// TIA Portal project "Project2" (V18)

(* hardware
DEVICE "S7-1500/ET200MP station_1"  S7-1500 station
   slot 0: "Rail_0"  Rack  6ES7 590-1***0-0AA0
   slot 1: "PLC_1"  CPU 1516-3 PN/DP  6ES7 516-3AN01-0AB0  V2.8
      slot 3: "CPU display_1"  6ES7591-1BA00-0AA0
      slot 32768: "PROFINET interface_1"  X1
         slot 32769: "Port_1"  X1 P1
         slot 32770: "Port_2"  X1 P2
      slot 33024: "PROFINET interface_2"  X2
         slot 33025: "Port_1"  X2 P1
      slot 33280: "DP interface_1"  X3
      slot 34817: "Virtual CP interface port_1"  Virtual CP interface port  Virtual CP interface port
DEVICE "GSD device_1"  GSD.Device.PN
   slot 0: "Rack"  Rack  V1.0
   slot 0: "IND360"  IND360 2 Block Format  MT-IND36XXXXXX  V1.0.0
      slot 0: "DAP 2 Block Parameter"  DAP 2 Block Parameter
      slot 1: "PROFINET"  PROFINET
         slot 1: "Port 1"  Port 1
         slot 2: "Port 2"  Port 2
      slot 1: "Measuring Block 1_1"  Measuring Block 1
         slot 0: "Parameter Access Point"  Parameter Access Point
         slot 1: "MB Command Value"  MB Command Value
         slot 2: "MB Channel Mask"  MB Channel Mask
         slot 3: "MB Command"  MB Command
         slot 4: "MB Measuring Value"  MB Measuring Value
         slot 5: "MB Device Status"  MB Device Status
         slot 6: "MB Response"  MB Response
      slot 2: "Status Block_1"  Status Block
         slot 0: "Parameter Access Point"  Parameter Access Point
         slot 1: "SB Reserved 1"  SB Reserved 1
         slot 2: "SB Reserved 2"  SB Reserved 2
         slot 3: "SB Reserved 3"  SB Reserved 3
         slot 4: "SB Command"  SB Command
         slot 5: "SB Status Group 1"  SB Status Group 1
         slot 6: "SB Status Group 2"  SB Status Group 2
         slot 7: "SB Status Group 3"  SB Status Group 3
         slot 8: "SB Response"  SB Response
DEVICE "HMI_1"  KTP400 Basic PN
   slot 0: "HMI_1"  KTP400 Basic PN  6AV2 123-2DB03-0AX0  17.0.0.0
   slot 1: "HMI_RT_1"  KTP400 Basic PN  6AV2 123-2DB03-0AX0  17.0.0.0
   slot 5: "HMI_1.IE_CP_1"  PROFINET Interface  17.0.0.0
      slot 1: "PROFINET Interface_1"  PROFINET Interface
         slot 1: "Port_1"  Port
*)

// ===== PLC "PLC_1"  CPU 1516-3 PN/DP =====

VAR_GLOBAL   // PLC tag table "Default tag table"
   "FirstScan" AT %M1.0 : Bool;
END_VAR

VAR_GLOBAL   // PLC tag table "IND"
   "T_MB_CmdValue" AT %QD0 : Real;
   "T_MB_Command" AT %QW6 : Word;
   "T_MB_Response" AT %IW6 : Word;
   "T_MB_Value" AT %ID0 : Real;
   "T_MB_DevStatus" AT %IW4 : Word;
   "T_SB_StaGroup1" AT %IW8 : Word;
   "T_SB_StaGroup2" AT %IW10 : Word;
   "T_SB_StaGroup3" AT %IW12 : Word;
   "T_SB_Response" AT %IW14 : Word;
   "T_SB_Command" AT %QW14 : Word;
   "AlibiGross_Byte(0)" AT %MB50 : Byte;
   "AlibiGross_Byte(1)" AT %MB51 : Byte;
   "AlibiGross_Byte(2)" AT %MB52 : Byte;
   "AlibiGross_Byte(3)" AT %MB53 : Byte;
   "AlibiNet_Byte(0)" AT %MB58 : Byte;
   "AlibiNet_Byte(1)" AT %MB59 : Byte;
   "AlibiNet_Byte(2)" AT %MB60 : Byte;
   "AlibiNet_Byte(3)" AT %MB61 : Byte;
   "AlibiTare_Byte(0)" AT %MB66 : Byte;
   "AlibiTare_Byte(1)" AT %MB67 : Byte;
   "AlibiTare_Byte(2)" AT %MB68 : Byte;
   "AlibiTare_Byte(3)" AT %MB69 : Byte;
   "AlibiGross_Real" AT %MD50 : Real;
   "AlibiNet_Real" AT %MD58 : Real;
   "AlibiTare_Real" AT %MD66 : Real;
END_VAR

TYPE "SAI_MB_DeviceStatus"
VERSION : 0.1
   STRUCT
      "Alternate weight unit" : Bool;
      "Run flat" : Bool;
      "Device specific bit 2" : Bool;
      "Device specific bit 3" : Bool;
      "Device specific bit 4" : Bool;
      "Device specific bit 5" : Bool;
      "Device specific bit 6" : Bool;
      "Device specific bit 7" : Bool;
      "Sequence bit 0" : Bool;
      "Sequence bit 1" : Bool;
      "Heart Beat" : Bool;
      "Data OK" : Bool;
      "Alarm Condition" : Bool;
      "Center of Zero" : Bool;
      Motion : Bool;
      "Net Mode" : Bool;
   END_STRUCT;
END_TYPE

TYPE "SAI_SB_RedAlert"
   STRUCT
      "Zero out of range" : Bool;
      "Symetry errors" : Bool;
      "LC Temperature out of normal temperature" : Bool;
      "Weights and measures failure" : Bool;
      "Foreign device detected" : Bool;
      "Test mode" : Bool;
      "LC temperature out of operatio" : Bool;
      "LC parameters block checksum error" : Bool;
      "Calibration error" : Bool;
      "Out of A/D range over/under" : Bool;
      "Checksu failure" : Bool;
      "Weight blocked" : Bool;
      "LC Missing" : Bool;
      "Customer-defined overload" : Bool;
      "Customer-defined underload" : Bool;
   END_STRUCT;
END_TYPE

TYPE "SAI_SB_Alarm"
   STRUCT
      "LC overload in operation range" : Bool;
      "LC Mix" : Bool;
      "Application defined 1" : Bool;
      "Application defined 2" : Bool;
      "Application defined 3" : Bool;
      "Application defined 4" : Bool;
      "Application defined 5" : Bool;
      "Application defined 7" : Bool;
      "Rate of change error" : Bool;
      "Communication error" : Bool;
      "Over / under voltage" : Bool;
      "Weight drift" : Bool;
      Breach : Bool;
      "Calibration expired" : Bool;
      "Over Current" : Bool;
      "LC overload in normal range" : Bool;
   END_STRUCT;
END_TYPE

DATA_BLOCK "SAI_Cyclic_CheckAlive_DB"   // DB1
{ S7_Optimized_Access := 'FALSE' }
VERSION : 0.1
// stored: InstanceOfName SAI_Cyclic_CheckAlive
"SAI_Cyclic_CheckAlive"
BEGIN
END_DATA_BLOCK

DATA_BLOCK "SAI_Cyclic_WeightProc_DB"   // DB2
{ S7_Optimized_Access := 'FALSE' }
VERSION : 0.1
// stored: InstanceOfName SAI_Cyclic_WeightProc
"SAI_Cyclic_WeightProc"
BEGIN
END_DATA_BLOCK

FUNCTION_BLOCK "SAI_Cyclic_CheckAlive"   // FB1, LAD
TITLE = Check HearBeat status bit and update the Alive bit
{ S7_Optimized_Access := 'FALSE' }
VERSION : 0.1
   VAR_INPUT
      MB_DevStatus : Word;
   END_VAR
   VAR_OUTPUT
      Alive : Bool;
      HeartBeat : Bool;
   END_VAR
   VAR
      PTrigHeart : Bool;
      NTrigHeart : Bool;
      bResetTimer : Bool;
      IEC_Timer : IEC_TIMER;
   END_VAR
   VAR_TEMP
      DevStatus : "SAI_MB_DeviceStatus";
   END_VAR
   VAR_TEMP   // added for the SCL form of the ladder/FBD networks
      _w1 : Bool;
      _w2 : Bool;
      _w3 : Bool;
   END_VAR
BEGIN

REGION Network 1: 复制设备状态到结构体 / Gets the cyclic device status - HeartBeat bit
   // Gets the cyclic device status - HeartBeat bit
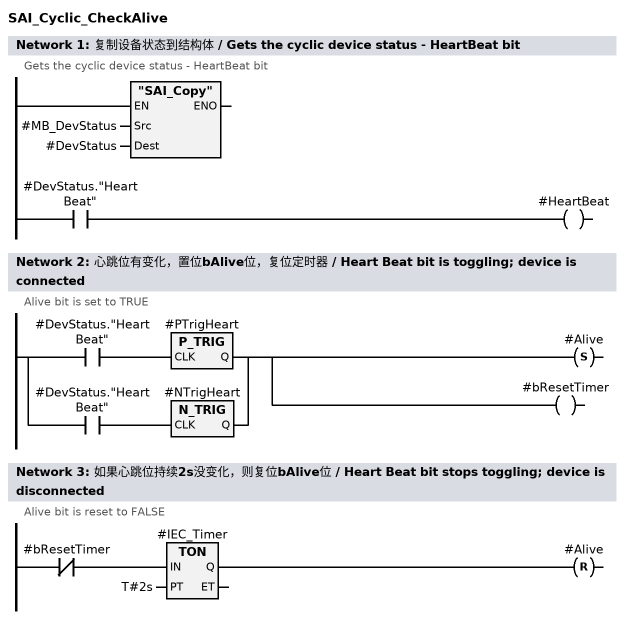
   RUNG wire#powerrail
      "SAI_Copy"(Src := #MB_DevStatus, Dest := #DevStatus)
   END_RUNG
   RUNG wire#powerrail
      Contact( #DevStatus."Heart Beat" )
      Coil( #HeartBeat )
   END_RUNG
   // the same network as SCL:
   "SAI_Copy"(Src := #MB_DevStatus, Dest := #DevStatus);
   #HeartBeat := #DevStatus."Heart Beat";
END_REGION

REGION Network 2: 心跳位有变化，置位bAlive位，复位定时器 / Heart Beat bit is toggling; device is connected
   // Alive bit is set to TRUE
   RUNG wire#powerrail
      Contact( #DevStatus."Heart Beat" )
      P_Trig( #PTrigHeart )
      wire#w1
      S_Coil( #Alive )
   END_RUNG
   RUNG wire#powerrail
      Contact( #DevStatus."Heart Beat" )
      N_Trig( #NTrigHeart )
   END_RUNG wire#w1
   RUNG wire#w1
      Coil( #bResetTimer )
   END_RUNG
   // the same network as SCL:
   #_w1 := #DevStatus."Heart Beat" AND NOT #PTrigHeart;   // rising edge
   #PTrigHeart := #DevStatus."Heart Beat";
   #_w2 := NOT #DevStatus."Heart Beat" AND #NTrigHeart;   // falling edge
   #NTrigHeart := #DevStatus."Heart Beat";
   #_w3 := #_w1 OR #_w2;
   IF #_w3 THEN #Alive := TRUE; END_IF;
   #bResetTimer := #_w3;
END_REGION

REGION Network 3: 如果心跳位持续2s没变化，则复位bAlive位 / Heart Beat bit stops toggling; device is disconnected
   // Alive bit is reset to FALSE
   #IEC_Timer.TON(IN := NOT #bResetTimer, PT := T#2s);
   IF #IEC_Timer.Q THEN #Alive := FALSE; END_IF;
END_REGION
END_FUNCTION_BLOCK

FUNCTION_BLOCK "SAI_Cyclic_WeightProc"   // FB2, LAD
TITLE = Cyclic Weighing Process: Send PLC commands and read Weight data and device status bits
{ S7_Optimized_Access := 'FALSE' }
VERSION : 0.1
   VAR_INPUT
      WeightCmd : Word := 3;
      MB_DevStatus : Word;
   END_VAR
   VAR_OUTPUT
      RealTimeWeight : Real;
      StableWeight : Real;
      DataOK : Bool;
      Motion : Bool;
      NetMode : Bool;
      Alarm : Bool;
      Done : Bool;
      Error : Bool;
   END_VAR
   VAR_IN_OUT
      TareImmediate : Bool;
      TareStable : Bool;
      ZeroImmediate : Bool;
      ZeroStable : Bool;
      PreTareValue : Real;
      PreTare : Bool;
      ClearTare : Bool;
      MB_Value : Real;
      MB_Response : Word;
      MB_CmdValue : Real;
      MB_Command : Word;
   END_VAR
   VAR
      WriteTrigger : Bool;
      RestoreTrigger : Bool;
      Cmd : Int;
      TareStablePTrigger : Bool;
      ZeroStablePTrigger : Bool;
      ZeroImmedTrigger : Bool;
      TareImmedTrigger : Bool;
      ClearTareTrigger : Bool;
      PreTareTrigger : Bool;
   END_VAR
   VAR_TEMP
      DevStatus : "SAI_MB_DeviceStatus";
   END_VAR
   VAR_TEMP   // added for the SCL form of the ladder/FBD networks
      _w1 : Bool;
   END_VAR
BEGIN

REGION Network 1: 第一次运行时，将默认重量命令赋值给循环区命令 / During 1st PLC scan, moves the default weight reporting command to the cyclic command output word
   // 第一次扫描，写入重量命令 / During 1st scan, moves the default weight reporting command to the cyclic command output word
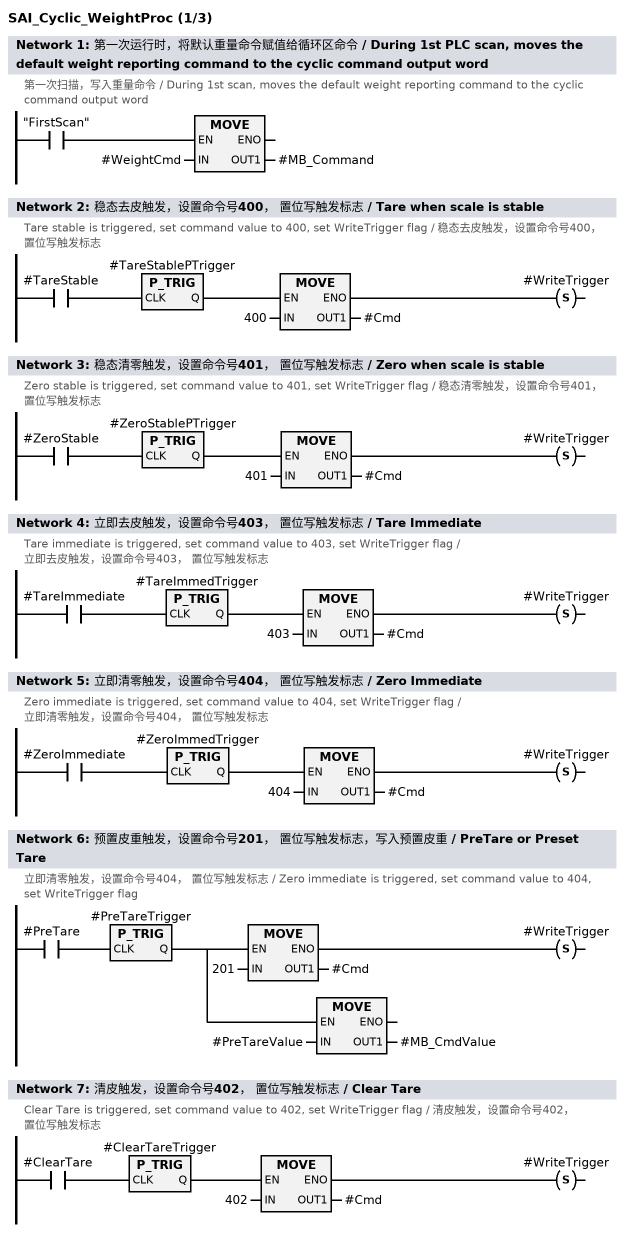
   RUNG wire#powerrail
      Contact( "FirstScan" )
      { S7_GenerateENO := "TRUE" } Move(in := #WeightCmd, out1 => #MB_Command)
   END_RUNG
   // the same network as SCL:
   IF "FirstScan" THEN #MB_Command := #WeightCmd; END_IF;
END_REGION

REGION Network 2: 稳态去皮触发，设置命令号400， 置位写触发标志 / Tare when scale is stable
   // Tare stable is triggered, set command value to 400, set WriteTrigger flag / 稳态去皮触发，设置命令号400， 置位写触发标志
   RUNG wire#powerrail
      Contact( #TareStable )
      P_Trig( #TareStablePTrigger )
      { S7_GenerateENO := "TRUE" } Move(in := 400, out1 => #Cmd)
      S_Coil( #WriteTrigger )
   END_RUNG
   // the same network as SCL:
   // ENO of a box is taken as its EN; it also drops when the box reports an error
   #_w1 := #TareStable AND NOT #TareStablePTrigger;   // rising edge
   #TareStablePTrigger := #TareStable;
   IF #_w1 THEN
       #Cmd := 400;
       #WriteTrigger := TRUE;
   END_IF;
END_REGION

REGION Network 3: 稳态清零触发，设置命令号401， 置位写触发标志 / Zero when scale is stable
   // Zero stable is triggered, set command value to 401, set WriteTrigger flag / 稳态清零触发，设置命令号401， 置位写触发标志
   RUNG wire#powerrail
      Contact( #ZeroStable )
      P_Trig( #ZeroStablePTrigger )
      { S7_GenerateENO := "TRUE" } Move(in := 401, out1 => #Cmd)
      S_Coil( #WriteTrigger )
   END_RUNG
   // the same network as SCL:
   // ENO of a box is taken as its EN; it also drops when the box reports an error
   #_w1 := #ZeroStable AND NOT #ZeroStablePTrigger;   // rising edge
   #ZeroStablePTrigger := #ZeroStable;
   IF #_w1 THEN
       #Cmd := 401;
       #WriteTrigger := TRUE;
   END_IF;
END_REGION

REGION Network 4: 立即去皮触发，设置命令号403， 置位写触发标志 / Tare Immediate
   // Tare immediate is triggered, set command value to 403, set WriteTrigger flag / 立即去皮触发，设置命令号403， 置位写触发标志
   RUNG wire#powerrail
      Contact( #TareImmediate )
      P_Trig( #TareImmedTrigger )
      { S7_GenerateENO := "TRUE" } Move(in := 403, out1 => #Cmd)
      S_Coil( #WriteTrigger )
   END_RUNG
   // the same network as SCL:
   // ENO of a box is taken as its EN; it also drops when the box reports an error
   #_w1 := #TareImmediate AND NOT #TareImmedTrigger;   // rising edge
   #TareImmedTrigger := #TareImmediate;
   IF #_w1 THEN
       #Cmd := 403;
       #WriteTrigger := TRUE;
   END_IF;
END_REGION

REGION Network 5: 立即清零触发，设置命令号404， 置位写触发标志 / Zero Immediate
   // Zero immediate is triggered, set command value to 404, set WriteTrigger flag / 立即清零触发，设置命令号404， 置位写触发标志
   RUNG wire#powerrail
      Contact( #ZeroImmediate )
      P_Trig( #ZeroImmedTrigger )
      { S7_GenerateENO := "TRUE" } Move(in := 404, out1 => #Cmd)
      S_Coil( #WriteTrigger )
   END_RUNG
   // the same network as SCL:
   // ENO of a box is taken as its EN; it also drops when the box reports an error
   #_w1 := #ZeroImmediate AND NOT #ZeroImmedTrigger;   // rising edge
   #ZeroImmedTrigger := #ZeroImmediate;
   IF #_w1 THEN
       #Cmd := 404;
       #WriteTrigger := TRUE;
   END_IF;
END_REGION

REGION Network 6: 预置皮重触发，设置命令号201， 置位写触发标志，写入预置皮重 / PreTare or Preset Tare
   // 立即清零触发，设置命令号404， 置位写触发标志 / Zero immediate is triggered, set command value to 404, set WriteTrigger flag
   RUNG wire#powerrail
      Contact( #PreTare )
      P_Trig( #PreTareTrigger )
      wire#w1
      { S7_GenerateENO := "TRUE" } Move(in := 201, out1 => #Cmd)
      S_Coil( #WriteTrigger )
   END_RUNG
   RUNG wire#w1
      { S7_GenerateENO := "TRUE" } Move(in := #PreTareValue, out1 => #MB_CmdValue)
   END_RUNG
   // the same network as SCL:
   // ENO of a box is taken as its EN; it also drops when the box reports an error
   #_w1 := #PreTare AND NOT #PreTareTrigger;   // rising edge
   #PreTareTrigger := #PreTare;
   IF #_w1 THEN
       #Cmd := 201;
       #WriteTrigger := TRUE;
       #MB_CmdValue := #PreTareValue;
   END_IF;
END_REGION

REGION Network 7: 清皮触发，设置命令号402， 置位写触发标志 / Clear Tare
   // Clear Tare is triggered, set command value to 402, set WriteTrigger flag / 清皮触发，设置命令号402， 置位写触发标志
   RUNG wire#powerrail
      Contact( #ClearTare )
      P_Trig( #ClearTareTrigger )
      { S7_GenerateENO := "TRUE" } Move(in := 402, out1 => #Cmd)
      S_Coil( #WriteTrigger )
   END_RUNG
   // the same network as SCL:
   // ENO of a box is taken as its EN; it also drops when the box reports an error
   #_w1 := #ClearTare AND NOT #ClearTareTrigger;   // rising edge
   #ClearTareTrigger := #ClearTare;
   IF #_w1 THEN
       #Cmd := 402;
       #WriteTrigger := TRUE;
   END_IF;
END_REGION

REGION Network 8: 将命令值赋值给输出循环区，复位标志，清除命令值 / Deliver the command
   // Move the command value to output, reset flags / 将命令输出，置位标志
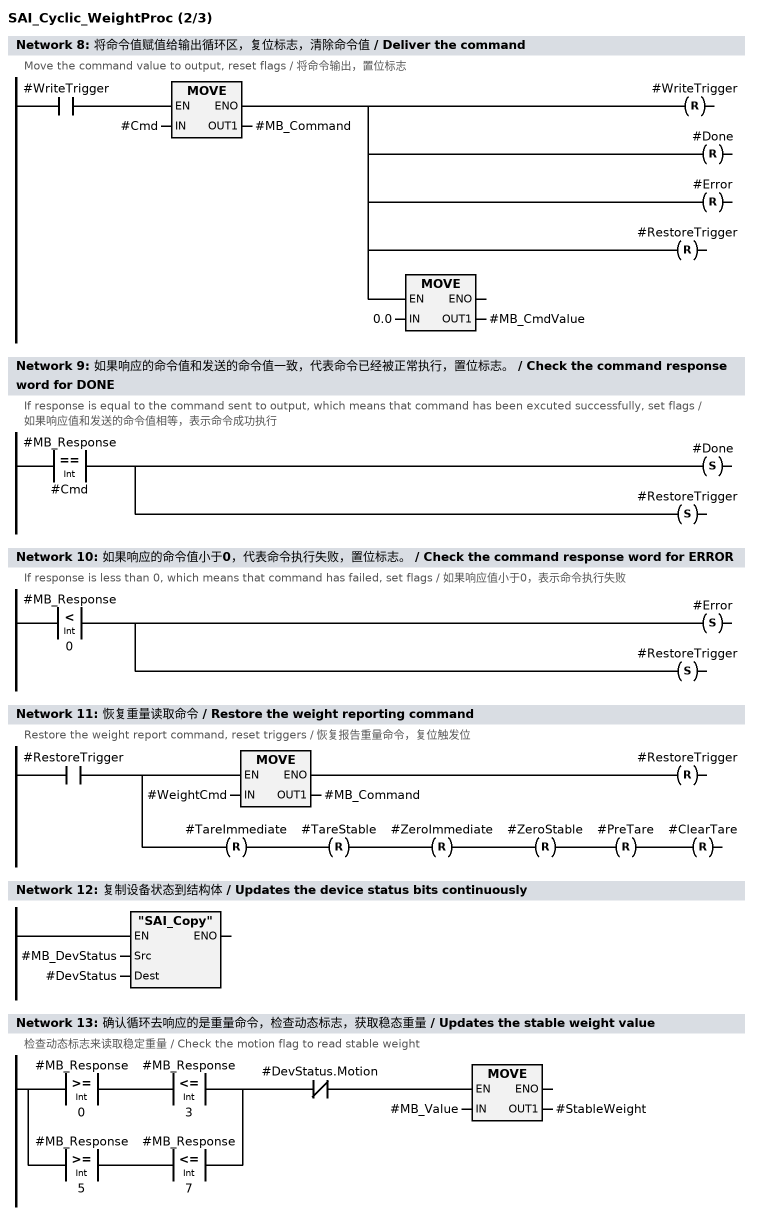
   RUNG wire#powerrail
      Contact( #WriteTrigger )
      { S7_GenerateENO := "TRUE" } Move(in := #Cmd, out1 => #MB_Command)
      wire#w1
      R_Coil( #WriteTrigger )
   END_RUNG
   RUNG wire#w1
      R_Coil( #Done )
   END_RUNG
   RUNG wire#w1
      R_Coil( #Error )
   END_RUNG
   RUNG wire#w1
      R_Coil( #RestoreTrigger )
   END_RUNG
   RUNG wire#w1
      { S7_GenerateENO := "TRUE" } Move(in := 0.0, out1 => #MB_CmdValue)
   END_RUNG
   // the same network as SCL:
   // ENO of a box is taken as its EN; it also drops when the box reports an error
   IF #WriteTrigger THEN #MB_Command := #Cmd; END_IF;
   #_w1 := #WriteTrigger;
   IF #_w1 THEN
       #WriteTrigger := FALSE;
       #Done := FALSE;
       #Error := FALSE;
       #RestoreTrigger := FALSE;
       #MB_CmdValue := 0.0;
   END_IF;
END_REGION

REGION Network 9: 如果响应的命令值和发送的命令值一致，代表命令已经被正常执行，置位标志。 / Check the command response word for DONE
   // If response is equal to the command sent to output, which means that command has been excuted successfully, set flags / 如果响应值和发送的命令值相等，表示命令成功执行
   RUNG wire#powerrail
      { S7_Templates := "SrcType := Int" } EQ_Contact(in1 := #MB_Response, in2 := #Cmd)
      wire#w1
      S_Coil( #Done )
   END_RUNG
   RUNG wire#w1
      S_Coil( #RestoreTrigger )
   END_RUNG
   // the same network as SCL:
   IF #MB_Response = #Cmd THEN
       #Done := TRUE;
       #RestoreTrigger := TRUE;
   END_IF;
END_REGION

REGION Network 10: 如果响应的命令值小于0，代表命令执行失败，置位标志。 / Check the command response word for ERROR
   // If response is less than 0, which means that command has failed, set flags / 如果响应值小于0，表示命令执行失败
   RUNG wire#powerrail
      { S7_Templates := "SrcType := Int" } LT_Contact(in1 := #MB_Response, in2 := 0)
      wire#w1
      S_Coil( #Error )
   END_RUNG
   RUNG wire#w1
      S_Coil( #RestoreTrigger )
   END_RUNG
   // the same network as SCL:
   IF #MB_Response < 0 THEN
       #Error := TRUE;
       #RestoreTrigger := TRUE;
   END_IF;
END_REGION

REGION Network 11: 恢复重量读取命令 / Restore the weight reporting command
   // Restore the weight report command, reset triggers / 恢复报告重量命令，复位触发位
   RUNG wire#powerrail
      Contact( #RestoreTrigger )
      wire#w1
      { S7_GenerateENO := "TRUE" } Move(in := #WeightCmd, out1 => #MB_Command)
      R_Coil( #RestoreTrigger )
   END_RUNG
   RUNG wire#w1
      R_Coil( #TareImmediate )
      R_Coil( #TareStable )
      R_Coil( #ZeroImmediate )
      R_Coil( #ZeroStable )
      R_Coil( #PreTare )
      R_Coil( #ClearTare )
   END_RUNG
   // the same network as SCL:
   // ENO of a box is taken as its EN; it also drops when the box reports an error
   IF #RestoreTrigger THEN #MB_Command := #WeightCmd; END_IF;
   #_w1 := #RestoreTrigger;
   IF #_w1 THEN
       #RestoreTrigger := FALSE;
       #TareImmediate := FALSE;
       #TareStable := FALSE;
       #ZeroImmediate := FALSE;
       #ZeroStable := FALSE;
       #PreTare := FALSE;
       #ClearTare := FALSE;
   END_IF;
END_REGION

REGION Network 12: 复制设备状态到结构体 / Updates the device status bits continuously
   RUNG wire#powerrail
      "SAI_Copy"(Src := #MB_DevStatus, Dest := #DevStatus)
   END_RUNG
   // the same network as SCL:
   "SAI_Copy"(Src := #MB_DevStatus, Dest := #DevStatus);
END_REGION

REGION Network 13: 确认循环去响应的是重量命令，检查动态标志，获取稳态重量 / Updates the stable weight value
   // 检查动态标志来读取稳定重量 / Check the motion flag to read stable weight
   RUNG wire#powerrail
      { S7_Templates := "SrcType := Int" } GE_Contact(in1 := #MB_Response, in2 := 0)
      { S7_Templates := "SrcType := Int" } LE_Contact(in1 := #MB_Response, in2 := 3)
      wire#w1
      I_Contact( #DevStatus.Motion )
      { S7_GenerateENO := "TRUE" } Move(in := #MB_Value, out1 => #StableWeight)
   END_RUNG
   RUNG wire#powerrail
      { S7_Templates := "SrcType := Int" } GE_Contact(in1 := #MB_Response, in2 := 5)
      { S7_Templates := "SrcType := Int" } LE_Contact(in1 := #MB_Response, in2 := 7)
   END_RUNG wire#w1
   // the same network as SCL:
   IF (((#MB_Response >= 0) AND (#MB_Response <= 3)) OR ((#MB_Response >= 5) AND (#MB_Response <= 7))) AND NOT #DevStatus.Motion THEN
       #StableWeight := #MB_Value;
   END_IF;
END_REGION

REGION Network 14: 确认循环去响应的是重量命令，读取实时的重量 / Updates the real time weight value
   // 读取实时重量 / Read real time weight
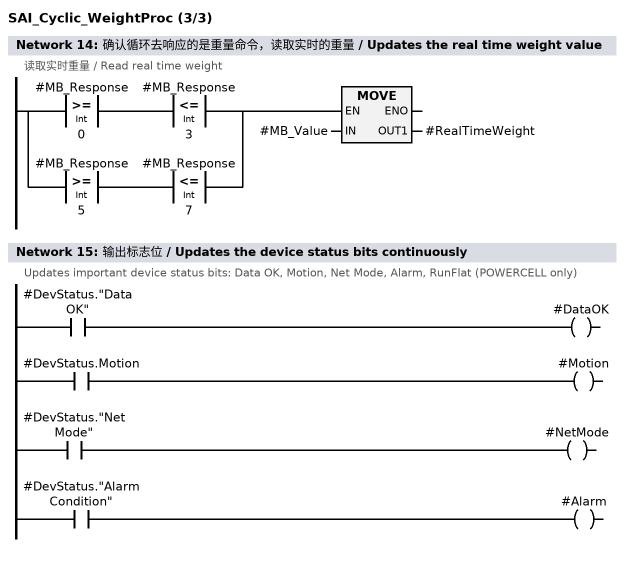
   RUNG wire#powerrail
      { S7_Templates := "SrcType := Int" } GE_Contact(in1 := #MB_Response, in2 := 0)
      { S7_Templates := "SrcType := Int" } LE_Contact(in1 := #MB_Response, in2 := 3)
      wire#w1
      { S7_GenerateENO := "TRUE" } Move(in := #MB_Value, out1 => #RealTimeWeight)
   END_RUNG
   RUNG wire#powerrail
      { S7_Templates := "SrcType := Int" } GE_Contact(in1 := #MB_Response, in2 := 5)
      { S7_Templates := "SrcType := Int" } LE_Contact(in1 := #MB_Response, in2 := 7)
   END_RUNG wire#w1
   // the same network as SCL:
   IF ((#MB_Response >= 0) AND (#MB_Response <= 3)) OR ((#MB_Response >= 5) AND (#MB_Response <= 7)) THEN
       #RealTimeWeight := #MB_Value;
   END_IF;
END_REGION

REGION Network 15: 输出标志位 / Updates the device status bits continuously
   // Updates important device status bits: Data OK, Motion, Net Mode, Alarm, RunFlat (POWERCELL only)
   RUNG wire#powerrail
      Contact( #DevStatus."Data OK" )
      Coil( #DataOK )
   END_RUNG
   RUNG wire#powerrail
      Contact( #DevStatus.Motion )
      Coil( #Motion )
   END_RUNG
   RUNG wire#powerrail
      Contact( #DevStatus."Net Mode" )
      Coil( #NetMode )
   END_RUNG
   RUNG wire#powerrail
      Contact( #DevStatus."Alarm Condition" )
      Coil( #Alarm )
   END_RUNG
   // the same network as SCL:
   #DataOK := #DevStatus."Data OK";
   #Motion := #DevStatus.Motion;
   #NetMode := #DevStatus."Net Mode";
   #Alarm := #DevStatus."Alarm Condition";
END_REGION
END_FUNCTION_BLOCK

FUNCTION "SAI_Copy" : Void   // FC1, LAD
{ S7_Optimized_Access := 'FALSE' }
VERSION : 0.1
   VAR_INPUT
      Src : Variant;
   END_VAR
   VAR_IN_OUT
      Dest : Variant;
   END_VAR
   VAR_TEMP
      TmpBuf : Array[0..100] of Byte;
      TmpRet : Int;
      TmpPos : DInt;
   END_VAR
BEGIN

REGION Network 1
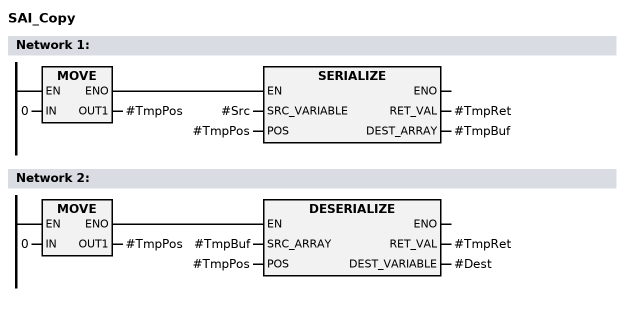
   // no SCL statement known for Serialize: written as a call
   #TmpPos := 0;
   #TmpRet := Serialize(SRC_VARIABLE := #Src, POS := #TmpPos, DEST_ARRAY => #TmpBuf);
END_REGION

REGION Network 2
   // no SCL statement known for Deserialize: written as a call
   #TmpPos := 0;
   #TmpRet := Deserialize(SRC_ARRAY := #TmpBuf, POS := #TmpPos, DEST_VARIABLE => #Dest);
END_REGION
END_FUNCTION

FUNCTION "MT_ACT_Application" : Void   // FC2, LAD
{ S7_Optimized_Access := 'FALSE' }
VERSION : 0.1
BEGIN

REGION Network 1: 循环重量处理 / Cyclic Weighing Data
   // 读取实时重量RealTimeWeight和稳态重量StableWeight，数据正常位DataOK，动态标志位Motion，净重模式位NetMode和警报位Alarm。
   // 上升沿触发执行稳态去皮TareStable，稳态清零ZeroStable，立即去皮TareImmediate，立即清零ZeroImmediate，预置皮重PreTare和清皮ClearTare，执行过程中，执行成功Done和失败Error的标志会复位为0，执行完成会置位Done或者Error来指示命令执行结果。清零去皮处理时，实时重量和稳态重量会保持不更新。
   // 在清零和去皮执行完成后，重量命令WeightCmd会自动发送一次，让MB Measuring Value循环区报告重量值，默认将恢复WeightCmd为读取净重（命令号3）。
   // 参照参数表中的重量命令值进行设置，执行清零或者去皮处理后，则会读取到对应的重量。
   // All the cyclical read and write commands can be issued from this Function Block.
   // The cyclic commands are triggered following a positive trigger. These commands are Tare Immediate, Tare Stable, Zero Immediate, Zero Stable, Pretare and Clear Tare. 
   // Upon successful execution of these commands, the DONE output bit will be set ON.
   // ERROR output bit will be set on if there is an error with the command execution.
   // Note: Only one cyclic command is possible at any one time.
   // If Net weight is required after executed a zero or tare command, insert decimal value "3" into the "WeightCmd" variable before triggering the cyclic scale command. Else, with decimal value "1" in the "WeightCmd" variable, the Function Block will return Gross Weight after the cyclic scale command. 
   // "DataOK" bit is set ON when the scale is in operation mode, not overloaded and not underload.
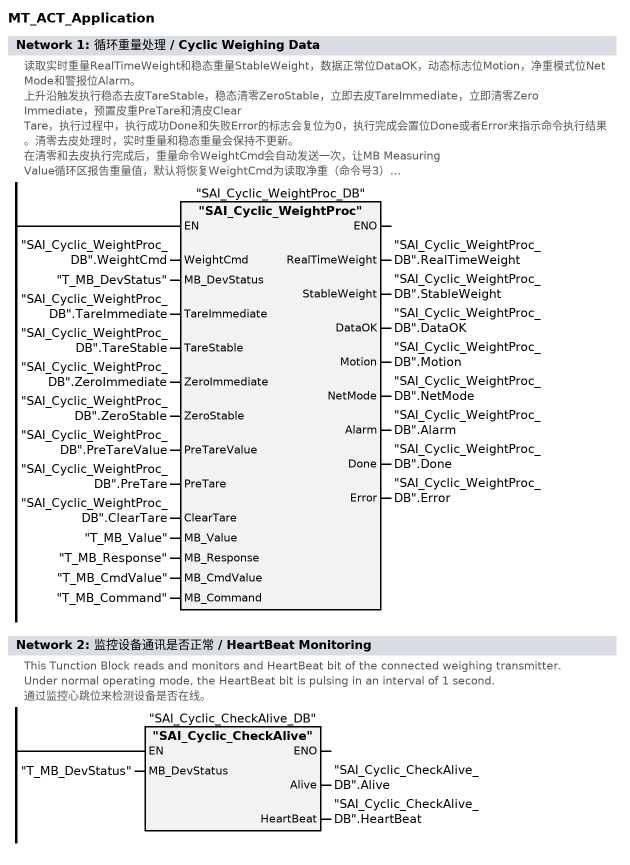
   RUNG wire#powerrail
      "SAI_Cyclic_WeightProc_DB"(WeightCmd := "SAI_Cyclic_WeightProc_DB".WeightCmd, MB_DevStatus := "T_MB_DevStatus", TareImmediate := "SAI_Cyclic_WeightProc_DB".TareImmediate, TareStable := "SAI_Cyclic_WeightProc_DB".TareStable, ZeroImmediate := "SAI_Cyclic_WeightProc_DB".ZeroImmediate, ZeroStable := "SAI_Cyclic_WeightProc_DB".ZeroStable, PreTareValue := "SAI_Cyclic_WeightProc_DB".PreTareValue, PreTare := "SAI_Cyclic_WeightProc_DB".PreTare, ClearTare := "SAI_Cyclic_WeightProc_DB".ClearTare, MB_Value := "T_MB_Value", MB_Response := "T_MB_Response", MB_CmdValue := "T_MB_CmdValue", MB_Command := "T_MB_Command", RealTimeWeight => "SAI_Cyclic_WeightProc_DB".RealTimeWeight, StableWeight => "SAI_Cyclic_WeightProc_DB".StableWeight, DataOK => "SAI_Cyclic_WeightProc_DB".DataOK, Motion => "SAI_Cyclic_WeightProc_DB".Motion, NetMode => "SAI_Cyclic_WeightProc_DB".NetMode, Alarm => "SAI_Cyclic_WeightProc_DB".Alarm, Done => "SAI_Cyclic_WeightProc_DB".Done, Error => "SAI_Cyclic_WeightProc_DB".Error)
   END_RUNG
   // the same network as SCL:
   "SAI_Cyclic_WeightProc_DB"(WeightCmd := "SAI_Cyclic_WeightProc_DB".WeightCmd,   // "SAI_Cyclic_WeightProc"
                           MB_DevStatus := "T_MB_DevStatus",
                           TareImmediate := "SAI_Cyclic_WeightProc_DB".TareImmediate,
                           TareStable := "SAI_Cyclic_WeightProc_DB".TareStable,
                           ZeroImmediate := "SAI_Cyclic_WeightProc_DB".ZeroImmediate,
                           ZeroStable := "SAI_Cyclic_WeightProc_DB".ZeroStable,
                           PreTareValue := "SAI_Cyclic_WeightProc_DB".PreTareValue,
                           PreTare := "SAI_Cyclic_WeightProc_DB".PreTare,
                           ClearTare := "SAI_Cyclic_WeightProc_DB".ClearTare,
                           MB_Value := "T_MB_Value",
                           MB_Response := "T_MB_Response",
                           MB_CmdValue := "T_MB_CmdValue",
                           MB_Command := "T_MB_Command",
                           RealTimeWeight => "SAI_Cyclic_WeightProc_DB".RealTimeWeight,
                           StableWeight => "SAI_Cyclic_WeightProc_DB".StableWeight,
                           DataOK => "SAI_Cyclic_WeightProc_DB".DataOK,
                           Motion => "SAI_Cyclic_WeightProc_DB".Motion,
                           NetMode => "SAI_Cyclic_WeightProc_DB".NetMode,
                           Alarm => "SAI_Cyclic_WeightProc_DB".Alarm,
                           Done => "SAI_Cyclic_WeightProc_DB".Done,
                           Error => "SAI_Cyclic_WeightProc_DB".Error);
END_REGION

REGION Network 2: 监控设备通讯是否正常 / HeartBeat Monitoring
   // This Tunction Block reads and monitors and HeartBeat bit of the connected weighing transmitter.
   // Under normal operating mode, the HeartBeat bit is pulsing in an interval of 1 second.
   // 通过监控心跳位来检测设备是否在线。
   RUNG wire#powerrail
      "SAI_Cyclic_CheckAlive_DB"(MB_DevStatus := "T_MB_DevStatus", Alive => "SAI_Cyclic_CheckAlive_DB".Alive, HeartBeat => "SAI_Cyclic_CheckAlive_DB".HeartBeat)
   END_RUNG
   // the same network as SCL:
   "SAI_Cyclic_CheckAlive_DB"(MB_DevStatus := "T_MB_DevStatus",   // "SAI_Cyclic_CheckAlive"
                           Alive => "SAI_Cyclic_CheckAlive_DB".Alive,
                           HeartBeat => "SAI_Cyclic_CheckAlive_DB".HeartBeat);
END_REGION
END_FUNCTION

ORGANIZATION_BLOCK "Main"   // OB1, LAD, ProgramCycle
TITLE = "Main Program Sweep (Cycle)"
{ S7_Optimized_Access := 'TRUE' }
VERSION : 0.1
   VAR_INPUT
      Initial_Call : Bool;   // Initial call of this OB
      Remanence : Bool;   // =True, if remanent data are available
   END_VAR
BEGIN

REGION Network 1
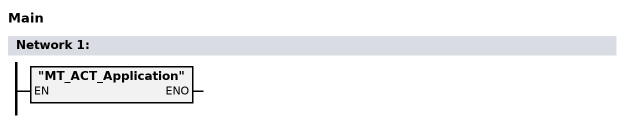
   RUNG wire#powerrail
      "MT_ACT_Application"()
   END_RUNG
   // the same network as SCL:
   "MT_ACT_Application"();
END_REGION
END_ORGANIZATION_BLOCK

(* ===== HMI "HMI_RT_1" =====
system functions are stored by id; their names below are inferred from use
connection "HMI_Connection_1": ETHERNET, SMART_S7_1500_OMS

HMI tags "Default tag table"
   "Tag_ScreenNumber" : UInt, internal
   "xHeartbeat" : Bool = PLC SAI_Cyclic_CheckAlive_DB.HeartBeat AT %DB1.DBX2.1, 1 s
   "rCurrentWeight" : Real = PLC SAI_Cyclic_WeightProc_DB.StableWeight AT %DB2.DBD8, 1 s
   "xZeroScale" : Bool = PLC SAI_Cyclic_WeightProc_DB.ZeroStable AT %DB2.DBX14.3, 1 s
   "xClearTare" : Bool = PLC SAI_Cyclic_WeightProc_DB.ClearTare AT %DB2.DBX20.1, 1 s
   "xSetTare" : Bool = PLC SAI_Cyclic_WeightProc_DB.TareStable AT %DB2.DBX14.1, 1 s

Template "Template_1" 480x272
   Button "Exit" at 388,227 size 63x44; TextOff 'Exit'; PictureOff "ExitRuntime_KTP400_Basic_PN_TR"; PictureOn "ExitRuntime_KTP400_Basic_PN_TR"
      on Release: StopRuntime(0)
   Button "Template_Button" at 268,227 size 63x44; TextOff 'Text'
   Button "Template_Button_1" at 148,227 size 63x44; TextOff 'Text'
   Button "Start screen" at 28,227 size 63x44; TextOff 'Start screen'; PictureOff "NavigateHome_KTP400_Basic_PN_TR"; PictureOn "NavigateHome_KTP400_Basic_PN_TR"
      on Release: ActivateScreen("Root screen", 0)
   SymbolicIOField "Symbolic_IO_Field_Screen" at 82,8 size 311x29; TextOff '0'; TextOn '1'; TextList "TextList_ScreenNames"
      ProcessValue <- "Tag_ScreenNumber"
      on Change: ActivateScreenByNumber("Tag_ScreenNumber", 0)
   DateTimeField "HmiScreenItemData" at 395,22 size 85x22
   DateTimeField "HmiScreenItemData_1" at 395,0 size 85x22
   GraphicView "Logo" at 0,0 size 80x45; Picture "Logo of HMI_1"

screen "Root screen" 480x272, template "Template_1"
   on GenerateScreen: SetTag("Tag_ScreenNumber", 1)
   TextField "HmiScreenItemData" at 42,58 size 100x30; Text 'IND360'
   TextField "Text field_1" at 57,98 size 90x25; Text 'Heartbeat'
   Rectangle "Rectangle_1" at 206,102 size 19x19
      Appearance <- "xHeartbeat"
   TextField "Text field_2" at 58,133 size 135x25; Text 'Current Weight'
   IOField "I/O field_1" at 206,130 size 68x32; FormatPattern s9.99; Unit  kg
      ProcessValue <- "rCurrentWeight"
   Button "Button_1" at 299,88 size 96x32; TextOff 'Zero Scale'
      on Press: function_b14e0dd5("xZeroScale", 0)
   Button "Button_2" at 299,126 size 96x32; TextOff 'Set Tare'
      on Press: function_b14e0dd5("xSetTare", 0)
   Button "Button_3" at 299,167 size 96x32; TextOff 'Clear Tare'
      on Press: function_b14e0dd5("xClearTare", 0)
*)